(* IEC 61131-3 sources: plc-vscode/tests/st/test-ready/trust-platform/examples/trust-twin/robot-cell/src, 2 files *)

(* ---- Robot_P3MinimalArm.fb.st ---- *)
(* trust-twin-generated: robot function block v1 *)
(* model: P3MinimalArm *)
(* manifest_hash: sha256:9236a9ea889aa5615171e7fc0bbadf3539e12216c5f7789639905366b7f63375 *)
(* urdf: crates/trust-runtime/tests/fixtures/p3_minimal_arm.urdf *)
(* base_frame: base, tool_frame: tool, grip_frame: workpiece.grip *)
(* joints: base_to_link_1->Joint1, link_1_to_link_2->Joint2 *)
(* native_bridge: trust_runtime::world::arm::step_robot_p3_minimal_arm_bridge *)
(* FK and URDF-derived poses are verified in trust_runtime::world::arm; this FB does not write transforms. *)

FUNCTION_BLOCK Robot_P3MinimalArm
VAR_INPUT
    Enable : BOOL;
    Command : INT;
END_VAR
VAR_OUTPUT
    EnabledOut : BOOL;
    Busy : BOOL;
    Done : BOOL;
    Fault : BOOL;
    State : INT;
    Owner : INT;
    HasWorkpiece : BOOL;
    GripperOpen : BOOL;
    StatusLight : BOOL;
    Joint1 : REAL;
    Joint2 : REAL;
    ToolYaw : REAL;
    ToolX : REAL;
    ToolY : REAL;
    ToolZ : REAL;
    WorkpieceX : REAL;
    WorkpieceY : REAL;
    WorkpieceZ : REAL;
END_VAR
END_FUNCTION_BLOCK

(* ---- main.st ---- *)
PROGRAM Main
VAR
    Robot : Robot_P3MinimalArm;
    RobotCommand : INT := 0;
    RobotMotionStep : INT := 0;
    RobotCycleTick : INT := 0;
    RobotShoulderAngle : REAL := -0.60;
    RobotElbowAngle : REAL := 0.35;
    RobotWristAngle : REAL := 0.25;
    RobotGripperOpen : BOOL := TRUE;
    RobotGripperX : REAL := 0.00;
    RobotGripperY : REAL := 0.80;
    RobotGripperZ : REAL := 0.00;
    RobotBoxX : REAL := 0.00;
    RobotBoxY : REAL := 0.35;
    RobotBoxZ : REAL := 0.00;
    RobotEnabled : BOOL := TRUE;
    RobotStatusLight : BOOL := FALSE;
END_VAR

RobotCycleTick := RobotCycleTick + 1;
IF RobotCycleTick >= 70 THEN
    RobotCycleTick := 0;
END_IF;

IF RobotCycleTick < 10 THEN
    (* approach pickup *)
    RobotCommand := 1;
ELSIF RobotCycleTick < 20 THEN
    (* close gripper *)
    RobotCommand := 2;
ELSIF RobotCycleTick < 30 THEN
    (* lift *)
    RobotCommand := 3;
ELSIF RobotCycleTick < 40 THEN
    (* translate *)
    RobotCommand := 4;
ELSIF RobotCycleTick < 50 THEN
    (* lower *)
    RobotCommand := 5;
ELSIF RobotCycleTick < 60 THEN
    (* open gripper *)
    RobotCommand := 6;
ELSE
    (* return *)
    RobotCommand := 7;
END_IF;

Robot(Enable := RobotEnabled, Command := RobotCommand);

RobotMotionStep := Robot.State;
RobotShoulderAngle := Robot.Joint1;
RobotElbowAngle := Robot.Joint2;
RobotWristAngle := Robot.ToolYaw;
RobotGripperOpen := Robot.GripperOpen;
RobotGripperX := Robot.ToolX;
RobotGripperY := Robot.ToolY;
RobotGripperZ := Robot.ToolZ;
RobotBoxX := Robot.WorkpieceX;
RobotBoxY := Robot.WorkpieceY;
RobotBoxZ := Robot.WorkpieceZ;
RobotEnabled := Robot.EnabledOut;
RobotStatusLight := Robot.StatusLight;
END_PROGRAM
